(* IEC 61131-3 sources: SortJet_MasterSPS_Aufbau.fbsproj/Device.device.xml.v3^/Plc Logic.plclogic.xml.v3^/Application.application.xml.v3^/09_Station/Stationen/Drehstation [207]/0_Konfig, 3 files *)

(* ---- Antriebsinformationen_207.gvl ---- *)
(* METADATA
{
	"v3Meta": {
		"objectGuid": "9d7b2ddc-bc65-44fc-9f07-0caa3fddbc7e"
	}
}
*)
{attribute 'allow_unqualified_access'}
NAMESPACE Antriebsinformationen_207
VAR_GLOBAL

//-------------------------------------------------------------------------------------------------
// ANTRIEBSINFORMATION [DREHSTATION]
//-------------------------------------------------------------------------------------------------

  apgInfoStation207Glastransport : ARRAY[cWAND_1..cANZAHL_WAENDE] OF AntriebsInformationen := [
    (
      wAchsID                                 :=     17,  // Achs ID aus dem EConSet
      stTyp                                   := 'Belt',  // Typ
      wpSchaltschrank                         :=   2040,  // Daten aus dem Schaltplan
      wpSchaltplanreihe                       :=     02,  // Daten aus dem Schaltplan
      wpSchaltplanseite                       :=    100,  // Daten aus dem Schaltplan
      rpMaxGeschwindigkeit                    :=   1000,  // [mm/s]   Max- Geschwindigkeit für den Automatikbetrieb
      rpHandGeschwindigkeit                   :=    200,  // [mm/s]   Hand- Geschwindigkeit
      rpReduzierteGeschwindigkeit             :=    67,   // [mm/s]   Reduzierte Geschwindigkeit
      rpReferenzGeschwindigkeit               :=      0,  // [mm/s]   Geschwindigkeit für die Referenzfahrt
      rpEinrichtGeschwindigkeit               :=     50,  // [mm/s]   Max Geschwindigkeit während der Einrichtung der Anlage
      rpMaxBeschleunigung                     :=   1500,  // [mm/s^2] Max Beschleunigung
      rpMaxVerzoegerung                       :=   2000,  // [mm/s^2] Max Verzoegerung
      rpMaxRuckzeit                           :=     50,  // [ms]     Ruckzeit des Antriebs
      rpReduzierteBeschleunigung              :=    500,  // [mm/s^2] Reduzierte Beschleunigung
      rpReduzierteVerzoegerung                :=    500,  // [mm/s^2] Reduzierte Verzoegerung
      rpBeschleunigungFremdanlage             :=   1000,  // [mm/s^2] Beschleunigung zu einer Fremdanlage
      rpGeschwindigkeitMessen                 :=    667,  // [mm/s] Geschwindigkeit beim Scheiben messen
      rpGeschwindigkeitSystemcheck            :=  500.0,  // [mm/s]   Geschwindigkeit im Systemcheck (nur Glastransport)
      rpGeschwindigkeitSystemcheckReduzierung :=  167.0,  // [mm/s]   Geschwindigkeit im Systemcheck bei belegtem Vorstop-Sensor (nur Glastransport)
      stOptionen                              := ( eEndschalterQuelle    := Endschalterquelle_EN.KEINE,     // Hardware-Endschalter: KEINE, UMRICHTER oder SPS
                                                   bVersorgungUeberXVR   := FALSE,                          // XVR-Modus: brueckt Hauptschalter 400 V und LS 230 V
                                                   bBremseLoesenFreigabe := FALSE )                         // Der Antrieb darf über eine Betriebsart die Bremse lösen
    )];

  apgInfoStation207GlastransportSlave : ARRAY[cWAND_1..cANZAHL_WAENDE] OF AntriebsInformationen := [
    (
      wAchsID                                 :=     65,  // Achs ID aus dem EConSet
      stTyp                                   := 'Belt',  // Typ
      wpSchaltschrank                         :=   2041,  // Daten aus dem Schaltplan
      wpSchaltplanreihe                       :=     02,  // Daten aus dem Schaltplan
      wpSchaltplanseite                       :=    100,  // Daten aus dem Schaltplan
      rpMaxGeschwindigkeit                    :=      0,  // [mm/s]   Max- Geschwindigkeit für den Automatikbetrieb
      rpHandGeschwindigkeit                   :=      0,  // [mm/s]   Hand- Geschwindigkeit
      rpReduzierteGeschwindigkeit             :=      0,  // [mm/s]   Reduzierte Geschwindigkeit
      rpReferenzGeschwindigkeit               :=      0,  // [mm/s]   Geschwindigkeit für die Referenzfahrt
      rpEinrichtGeschwindigkeit               :=      0,  // [mm/s]   Max Geschwindigkeit während der Einrichtung der Anlage
      rpMaxBeschleunigung                     :=      0,  // [mm/s^2] Max Beschleunigung
      rpMaxVerzoegerung                       :=      0,  // [mm/s^2] Max Verzoegerung
      rpMaxRuckzeit                           :=      0,  // [ms]     Ruckzeit des Antriebs
      rpReduzierteBeschleunigung              :=      0,  // [mm/s^2] Reduzierte Beschleunigung
      rpReduzierteVerzoegerung                :=      0,  // [mm/s^2] Reduzierte Verzoegerung
      rpBeschleunigungFremdanlage             :=      0,  // [mm/s^2] Beschleunigung zu einer Fremdanlage
      rpGeschwindigkeitMessen                 :=      0,  // [mm/s] Geschwindigkeit beim Scheiben messen
      rpGeschwindigkeitSystemcheck            :=  500.0,  // [mm/s]   Geschwindigkeit im Systemcheck (nur Glastransport)
      rpGeschwindigkeitSystemcheckReduzierung :=  167.0,  // [mm/s]   Geschwindigkeit im Systemcheck bei belegtem Vorstop-Sensor (nur Glastransport)
      stOptionen                              := ( eEndschalterQuelle    := Endschalterquelle_EN.KEINE,     // Hardware-Endschalter: KEINE, UMRICHTER oder SPS
                                                   bVersorgungUeberXVR   := FALSE,                          // XVR-Modus: brueckt Hauptschalter 400 V und LS 230 V
                                                   bBremseLoesenFreigabe := FALSE )                         // Der Antrieb darf über eine Betriebsart die Bremse lösen
    )];

  apgInfoStation207Drehen : AntriebsInformationen :=
    (
      wAchsID                                 :=        18,  // Achs ID aus dem EConSet
      stTyp                                   := 'Turning',  // Typ
      wpSchaltschrank                         :=      2042,  // Daten aus dem Schaltplan
      wpSchaltplanreihe                       :=        02,  // Daten aus dem Schaltplan
      wpSchaltplanseite                       :=        65,  // Daten aus dem Schaltplan
      rpMaxGeschwindigkeit                    :=       350,  // [Grad/s] MAX- Geschwindigkeit für die der Antrieb ausgelegt ist // Max 556
      rpHandGeschwindigkeit                   :=       150,  // [Grad/s] Hand- Geschwindigkeit
      rpReduzierteGeschwindigkeit             :=        20,  // [Grad/s] Reduzierte Geschwindigkeit für die bestimmte Situationen
      rpReferenzGeschwindigkeit               :=         1,  // [Grad/s] Geschwindigkeit für die Referenzfahrt
      rpEinrichtGeschwindigkeit               :=        10,  // [Grad/s] Max Geschwindigkeit während der Einrichtung der Anlage
      rpMaxBeschleunigung                     :=       300,  // [Grad/s^2] max Beschleunigung für die der Antrieb ausgelegt ist // Max 1026
      rpMaxVerzoegerung                       :=       300,  // [Grad/s^2] max Verzoegerung für die der Antrieb ausgelegt ist // Max 1026
      rpMaxRuckzeit                           :=       200,   // [ms]     Ruckzeit des Antriebs
      rpReduzierteBeschleunigung              :=       0.5,  // [Grad/s^2] Reduzierte Beschleunigung
      rpReduzierteVerzoegerung                :=       0.5,  // [Grad/s^2] Reduzierte Verzoegerung
      rpBeschleunigungFremdanlage             :=       0.5,  // [Grad/s^2] Beschleunigung zu einer Fremd-Anlage
      rpGeschwindigkeitMessen                 :=         0,  // [Grad/s] Geschwindigkeit für die Messfahrt
      rpGeschwindigkeitSystemcheck            :=  500.0,  // [mm/s]   Geschwindigkeit im Systemcheck (nur Glastransport)
      rpGeschwindigkeitSystemcheckReduzierung :=  167.0,  // [mm/s]   Geschwindigkeit im Systemcheck bei belegtem Vorstop-Sensor (nur Glastransport)
      stOptionen                              := ( eEndschalterQuelle    := Endschalterquelle_EN.UMRICHTER, // Hardware-Endschalter: KEINE, UMRICHTER oder SPS
                                                   bVersorgungUeberXVR   := FALSE,                          // XVR-Modus: brueckt Hauptschalter 400 V und LS 230 V
                                                   bBremseLoesenFreigabe := FALSE )                         // Der Antrieb darf über eine Betriebsart die Bremse lösen
    );

  apgInfoStation207Kippen : AntriebsInformationen :=
    (
      wAchsID                                 :=        65,  // Achs ID aus dem EConSet
      stTyp                                   := 'Tilting',  // Typ
      wpSchaltschrank                         :=      2043,  // Daten aus dem Schaltplan
      wpSchaltplanreihe                       :=         2,  // Daten aus dem Schaltplan
      wpSchaltplanseite                       :=       100,  // Daten aus dem Schaltplan
      rpMaxGeschwindigkeit                    :=      1400,  // [Grad/s] Max- Geschwindigkeit für die der Antrieb ausgelegt ist
      rpHandGeschwindigkeit                   :=      1400,  // [Grad/s] Hand- Geschwindigkeit
      rpReduzierteGeschwindigkeit             :=       800,  // [Grad/s] Reduzierte Geschwindigkeit für die bestimmte Situationen
      rpReferenzGeschwindigkeit               :=       100,  // [Grad/s] Geschwindigkeit für die Referenzfahrt
      rpEinrichtGeschwindigkeit               :=       100,  // [Grad/s] Max Geschwindigkeit während der Einrichtung der Anlage
      rpMaxBeschleunigung                     :=       250,  // [Grad/s^2] Max Beschleunigung für die der Antrieb ausgelegt ist
      rpMaxVerzoegerung                       :=       250,  // [Grad/s^2] Max Verzoegerung für die der Antrieb ausgelegt ist
      rpMaxRuckzeit                           :=        50,  // [ms] Ruckzeit des Antriebs
      rpReduzierteBeschleunigung              :=       100,  // [Grad/s^2] Reduzierte Beschleunigung
      rpReduzierteVerzoegerung                :=       100,  // [Grad/s^2] Reduzierte Verzoegerung
      rpBeschleunigungFremdanlage             :=         1,  // [Grad/s^2] Beschleunigung zu einer Fremd-Anlage
      rpGeschwindigkeitMessen                 :=         0,  // [Grad/s] Geschwindigkeit für die Messfahrt
      rpGeschwindigkeitSystemcheck            := 500.0,  // [mm/s]   Geschwindigkeit im Systemcheck (nur Glastransport)
      rpGeschwindigkeitSystemcheckReduzierung := 167.0,  // [mm/s]   Geschwindigkeit im Systemcheck bei belegtem Vorstop-Sensor (nur Glastransport)
      stOptionen                              := ( eEndschalterQuelle    := Endschalterquelle_EN.UMRICHTER, // Hardware-Endschalter: KEINE, UMRICHTER oder SPS
                                                   bVersorgungUeberXVR   := FALSE,                          // XVR-Modus: brueckt Hauptschalter 400 V und LS 230 V
                                                   bBremseLoesenFreigabe := FALSE )                         // Der Antrieb darf über eine Betriebsart die Bremse lösen
    );

    apgInfoStation207Querfahrt : AntriebsInformationen :=
    (
      wAchsID                                 :=         65,  // Achs ID aus dem EConSet
      stTyp                                   := 'Movement',  // Typ
      wpSchaltschrank                         :=       2044,  // Daten aus dem Schaltplan
      wpSchaltplanreihe                       :=         02,  // Daten aus dem Schaltplan
      wpSchaltplanseite                       :=        100,  // Daten aus dem Schaltplan
      rpMaxGeschwindigkeit                    :=        250,  // [mm/s] MAX- Geschwindigkeit für die der Antrieb ausgelegt ist
      rpHandGeschwindigkeit                   :=        100,  // [mm/s] Hand- Geschwindigkeit
      rpReduzierteGeschwindigkeit             :=         50,  // [mm/s] Reduzierte Geschwindigkeit für die bestimmte Situationen
      rpReferenzGeschwindigkeit               :=         20,  // [mm/s] Geschwindigkeit für die Referenzfahrt
      rpEinrichtGeschwindigkeit               :=         50,  // [mm/s] Max Geschwindigkeit während der Einrichtung der Anlage
      rpMaxBeschleunigung                     :=        600,  // [mm/s^2] max Beschleunigung für die der Antrieb ausgelegt ist
      rpMaxVerzoegerung                       :=        600,  // [mm/s^2] max Verzoegerung für die der Antrieb ausgelegt ist
      rpMaxRuckzeit                           :=        600,  // [ms]     Ruckzeit des Antriebs
      rpReduzierteBeschleunigung              :=        200,  // [mm/s^2] Reduzierte Beschleunigung
      rpReduzierteVerzoegerung                :=        200,  // [mm/s^2] Reduzierte Verzoegerung
      rpBeschleunigungFremdanlage             :=          0,  // [mm/s^2] Beschleunigung zu einer Fremd-Anlage
      rpGeschwindigkeitMessen                 :=          0,  // [mm/s] Geschwindigkeit für die Messfahrt
      rpGeschwindigkeitSystemcheck            := 500.0,  // [mm/s]   Geschwindigkeit im Systemcheck (nur Glastransport)
      rpGeschwindigkeitSystemcheckReduzierung := 167.0,  // [mm/s]   Geschwindigkeit im Systemcheck bei belegtem Vorstop-Sensor (nur Glastransport)
      stOptionen                              := ( eEndschalterQuelle    := Endschalterquelle_EN.UMRICHTER, // Hardware-Endschalter: KEINE, UMRICHTER oder SPS
                                                   bVersorgungUeberXVR   := FALSE,                          // XVR-Modus: brueckt Hauptschalter 400 V und LS 230 V
                                                   bBremseLoesenFreigabe := FALSE )                         // Der Antrieb darf über eine Betriebsart die Bremse lösen
    );

END_VAR

END_NAMESPACE

(* ---- MK_Station_207.gvl ---- *)
(* METADATA
{
	"v3Meta": {
		"objectGuid": "ad0b4350-ba92-412a-9245-7792853cbecb"
	}
}
*)
{attribute 'allow_unqualified_access'}
NAMESPACE MK_Station_207
VAR_GLOBAL

//-------------------------------------------------------------------------------------------------
// MASCHINEPARAMETER: DREHSTATION
//-------------------------------------------------------------------------------------------------

  apgMKStation207 : Parameter_Station:=
    (
      stStationsNummern                     := ( NummerIntern :=   207,                                                      // Stationsnummer fuer das MMI und die Stationsangabe der Meldungen
                                                 NummerExtern :=  1207,                                                      // Stationsnummer fuer Bedienermeldungen
                                                 NummerSPS    :=   207 ),                                                    // Stationsnummer SPS-intern (Indizes)
      bDeaktivieren                         := FALSE,                                                                        // Station deaktiviert (keine Auftraege, keine Referenzfahrt)
      wMeldungsNummer                       := 1810,                                                                         // Basis-Meldungsnummer (WatchIO)
      eStationsTyp                          := eStation,                                                                     // Typ der Station
      eaAutomatikkreis                      := [eAutomatikkreis_1],                                                          // Automatikkreise, zu denen die Station gehoert
      eaSicherheitskreis                    := [eSicherheitskreis_1, eSicherheitskreis_4],                                   // Sicherheitskreise, in die die Station eingebunden ist
      astSicherheitskreisTeilabschaltung    := [ ( eSicherheitskreis := eSicherheitskreis_4,                                 // SK4 (Abschrankung 208) schaltet nur Drehen/Kippen ab,
                                                   bTeilabschaltung  := TRUE,                                                //   Glastransport, Geblaese, Querfahrt und Pneumatik bleiben aktiv
                                                   bDrehen           := TRUE,
                                                   bKippen           := TRUE ) ],
      eSystemcheckZyklus                    := eSystemcheckZyklus_1,                                                         // In welchem Zyklus des Systemchecks die Station geprueft wird
      stSchnittstellendaten                 := ( wVorgaengerStation := cSTATION_DYNAMISCH,                                   // Station vor dieser Station (cSTATION_DYNAMISCH bei mehreren)
                                                 wNachfolgerStation := cSTATION_DYNAMISCH,                                   // Station nach dieser Station (cSTATION_DYNAMISCH bei mehreren)
                                                 bStationIstShuttle := FALSE                                                 // Station ist ein Shuttle
                                               ),
      stStationsOptionen                    := ( stSystemcheck :=  ( bScheibenVermessenSystemCheck               := TRUE,    // Scheiben im Systemcheck vermessen
                                                                     bScheibeNachSystemcheckAufAuslauf           := TRUE,    // Scheibe nach dem Systemcheck auf den Auslaufsensor fahren
                                                                     bSystemCheckMitVorgaengerBatchTransport     := FALSE,   // derzeit ohne Funktion
                                                                     bSystemCheckMitNachfolgerBatchTransport     := FALSE,   // derzeit ohne Funktion
                                                                     bOptionSystemCheckScheibeMittigLegen        := FALSE ), // derzeit ohne Funktion

                                                 // stTransfershuttle
                                                 stGlastransport :=  ( bVortransport                             := FALSE,   // Vortransport aktivieren [Bsp.: Nach einem Eintransport mit gesetztem Bit <Letzte Scheibe>]
                                                                       bTransportMasterSlaveEintransport         := FALSE,   // derzeit ohne Funktion
                                                                       bTransportMasterSlaveAustransport         := TRUE ,   // Austransport als Slave auf die Achse des Nachfolgers
                                                                       bGLasUebernahmeSenkrecht                  := FALSE,   // RKT - Eintransport in Senkrechter-Position bzw. in Waagerechter- Position [default]
                                                                       bAustransportISOLinie                     := FALSE,   // Austransport an eine ISO-Linie
                                                                       bScheibenVermessen                        := FALSE,   // Scheibenmessung am Anlegetisch/Anlegewand
                                                                       bMessrichtungNegativ                      := FALSE,   // Negative Fahrtrichtung beim Messen
                                                                       bScheibenmessungEintransport              := FALSE,   // Scheibenmessung beim Eintransport
                                                                       bScheibenmessungSensorVorabAuslauf        := FALSE    // Scheibenmessung mit SensorVorabAuslauf z.B. Anlegewand
                                                                      ),
                                                 // stAnlegetisch
                                                 // stEckuebergabe
                                                 stDrehstation   :=  ( bDrehpositionenVomMMI                     := FALSE,            // TRUE: Drehpositionen aus den MMI-Auftragsdaten; FALSE: aus der Stationskonfiguration [aEintransporte/aAustransporte]
                                                                       wStandardTransferstation                  := cSTATION_206 ),   // Systemcheck (Drehpositionen nicht vom MMI): Transferstation, wenn die Auftragsdaten 0 enthalten
                                                 bVorAbKomponentenAnsteuerung              := FALSE,                         // VorAbKomponentenAnsteuerung Auftraege werden bearbeitet
                                                 bVerstellungEinAusGefahrenLogikDrehen     := FALSE,                         // Verstellung: Logik ein-/ausgefahren gedreht
                                                 bLangsamfahrtNockenQuerfahrtAktivieren    := FALSE,                         // Querfahrt: Langsamfahrt-Nocken auswerten
                                                 bSKBlockierenDurchVorabSensoren           := FALSE,                         // Vorab-Sensoren belegt blockieren das Oeffnen des Sicherheitskreises
                                                 bStationLeerfahrenBeiSkAnforderung        := FALSE,                         // Station bei Anforderung Sicherheitskreis leerfahren
                                                 bGlasAbgenommenAutomatischQuittieren      := FALSE,                         // derzeit ohne Funktion
                                                 bScheibeAbnehmenNachEintransport          := FALSE                          // Scheibe nach dem Eintransport wieder abnehmen
                                               ),
      stStationsAufbau                      := ( bGeblase                      := [ cANZAHL_WAENDE(TRUE) ],                  // Ausbaustufe: Geblaese je Wand
                                                 bGlastransport                := [ cANZAHL_WAENDE(TRUE) ],                  // Ausbaustufe: Glastransport je Wand
                                                 bKippen                       := [ cANZAHL_WAENDE(TRUE) ],                  // Ausbaustufe: Kippen je Wand
                                                 bKippenSchuetz                := TRUE,                                      // Kippen ueber Schuetz statt Umrichter
                                                 bTransportVerstellung         := [ cANZAHL_WAENDE(FALSE) ],                 // Ausbaustufe Shuttle: Transport-/Dickenverstellung je Wand
                                                 bHub                          := FALSE,                                     // Ausbaustufe: Hub der Station
                                                 bHubrahmen                    := FALSE,                                     // Ausbaustufe: Hubrahmen (Riemen heben/senken)
                                                 bDrehen                       := TRUE,                                      // Ausbaustufe: Drehen
                                                 bQuerachse                    := FALSE,                                     // Ausbaustufe: Querachse
                                                 bMessachse                    := FALSE,                                     // Ausbaustufe: Messachse (Anlegetisch, Anlegewand)
                                                 bDruckluft                    := TRUE,                                      // Druckluftueberwachung vorhanden
                                                 bAnschlag                     := FALSE,                                     // Ausbaustufe: Ausrichtanschlaege
                                                 bSensorAuslauf                := TRUE,                                      // Auslaufsensor vorhanden
                                                 bSensorEinlauf                := TRUE,                                      // Einlaufsensor vorhanden
                                                 bSensorEinlaufStopp           := FALSE,                                     // Shuttle: zusaetzlicher Stopp-Sensor am Einlauf (ohne: Einlaufsensor), Gegenstueck zum Auslauf-Stopp im Rueckwaertstransport
                                                 bSensorAuslaufStopp           := FALSE,                                     // Shuttle: zusaetzlicher Stopp-Sensor am Auslauf (ohne: Auslaufsensor), Verfahrfreigabe und Scheibe hat Shuttle verlassen
                                                 bDurchlaufSperreZumNachfolger := FALSE,                                     // Ausbaustufe: bewegliche Abschrankung zum Nachfolger
                                                 bQuerfahrt                    := FALSE,                                     // Ausbaustufe: Querfahrt
                                                 bKipparme                     := FALSE,                                     // Ausbaustufe: Kipparme
                                                 bSlaveAntrieb                 := FALSE,                                     // Glastransport mit Slave-Antrieb
                                                 bMessachseAmEndeVomTisch      := FALSE,                                     // Messachse am Ende des Tisches (Hoehenfehler fragt den Bediener)
                                                 bWandverstellung              := [ FALSE ],                                 // Ausbaustufe Station: Wandverstellung je Wand
                                                 bWandverstellungMotorisch     := FALSE,                                     // Shuttle: Transport-/Wandverstellung mit Antrieb statt pneumatisch
                                                 bRoellchenleiste              := [ FALSE ],                                 // Ausbaustufe Station: Roellchenleiste je Wand
                                                 bDurchgang                    := FALSE,                                     // Station ist Teil eines Durchgangs (belegt = Oeffnen blockiert)
                                                 bRolltor                      := FALSE,                                     // Ausbaustufe Faecherwagen: Rolltor
                                                 bKlemmzylinder                := FALSE,                                     // Ausbaustufe Faecherwagen: Klemmzylinder fixiert den Oberrahmen beim Ein- und Ausschleusen
                                                 bGreifer                      := [cANZAHL_WAENDE(FALSE)],                   // Shuttle: Greifer je Wand (Scheibe aus dem Faecherwagen ziehen bzw. hineinschieben)
                                                 bRFID                         := FALSE,                                     // RFID-Leser vorhanden
                                                 bAGV                          := FALSE,                                     // Ausbaustufe Faecherwagen: Betrieb mit AGV
                                                 bDLSSchmiersystem             := FALSE,                                     // Zentralschmierung DLS vorhanden
                                                 bGlastransportSlaveVorhanden  := FALSE,                                     // Glastransport mit Slave-Antrieb (Meldungen/Ueberwachung Slave)
                                                 wHydraulikstation             := 0                                          // Faecherwagen Hydraulik: zugeordnete Hydraulikstation (cHYDRAULIKSTATION_x), 0 = keine
                                               ),
      stStationsParameter                   := ( rLaengeUebergroesseScheibe              := 4240,                            // Shuttle: ab dieser Scheibenlaenge gilt die Scheibe als uebergross [mm]
                                                 rMinGlasHoeheAutomatischenEintransport  := 500,                             // VSG: Mindesthoehe fuer automatischen Eintransport [mm]
                                                 rMinGlasLaengeAutomatischenEintransport := 500,                             // VSG: Mindestlaenge fuer automatischen Eintransport [mm]
                                                 wMaximaleAnzahlAktiverAuftraege := 1,                                       // derzeit ohne Funktion
                                                 rMinPosSwEsEingrenzung                  := 0.0,                             // Externer zusaetzlicher Software-Endschalter MIN; 0 = inaktiv; darf den MK-MIN nur weiter eingrenzen
                                                 rMaxPosSwEsEingrenzung                  := 0.0,                             // Externer zusaetzlicher Software-Endschalter MAX; 0 = inaktiv; darf den MK-MAX nur weiter eingrenzen
                                                 rPosFreigabePufferAusfahren             := 0.0                              // derzeit ohne Funktion
                                              ),
      // stFremdanlage
      stGlasdaten                           := [(
                                                 rlMinGlasLaenge                  := 350,                                    // minimal zulässige GlasLänge
                                                 rlMaxGlasLaenge                  := 2500,                                   // maximale zulässige GlasLänge
                                                 rlMinGlasHoehe                   := 190,                                    // minimal zulässige GlasHöhe
                                                 rlMaxGlasHoehe                   := 1800,                                   // maximale zulässige GlasHöhe
                                                 rlMinGlasDicke                  := 3,                                     // minimal zulässige GlasDicke
                                                 rlMaxGlasDicke                  := 12.76,                                      // maximal zulaessige Glasdicke [mm]
                                                 rlLaengeMaxGlas                  := 0.0                                     // maximal zulaessige Glaslaenge [mm]
                                               )]
      // astShuttleAnhaltenQuellen
    );

  apgMKStation207Glastransport : ARRAY[cWAND_1..cANZAHL_WAENDE] OF Parameter_Glastransport := [
    (
      rLaengeStation                        := 2800, // Länge der Station
      rScheibenabstand                      :=  300, // Der Abstand zwischen zwei Scheiben auf der Station
      rWegUeberAuslauf                      :=   50, // Weg ueber den Auslaufsensor hinaus [mm]
      rWegUeberEinlauf                      :=   50, // Weg ueber den Einlaufsensor hinaus [mm]
      rWegUeberSensorenSystemCheck          :=   15, // Der Weg der Ueber ein die Sensoren zum vermessen der Scheiben
      rUeberwachungAuslaufsensor            :=  500, // Ueberwachung des Auslaufsensors [Strecke in der der Auslaufsensor Frei / ueberfahren werden soll]
      rUeberwachungEinlaufsensor            :=  500, // Ueberwachung des Einlaufsensors [Strecke in der der Einlaufsensor Frei / ueberfahren werden soll]
      rWegUeberEinlaufEintransport          :=  150, // Eintransport vorwaerts: Abstand Scheibenhinterkante zum Einlaufsensor [mm]
      rWegUeberEinlaufAustransport          :=   50, // Lage Auf Einlauf: Scheibe liegt um diesen Weg auf dem Einlaufsensor [mm]
      rWegUeberAuslaufEintransport          :=   50, // Eintransport rueckwaerts: Abstand Scheibenhinterkante zum Auslaufsensor [mm]
      rWegUeberAuslaufAustransport          :=   10, // Lage Auf Auslauf: Weg ueber den Auslaufsensor hinaus [mm]
      rWegEinlaufsensorZuVorStopSensor      := 2700, // Beschreibt den Weg vum eine Scheibe beim EIntransport vom Einlaufsensor bis ueberden Vorabstopsensor zu verfahren
      rMesstoleranz                         :=   10, // Toleranz-Mass fuer die Scheibenlaengenmessung
      rMessstrecke                          := 2740, // Beschreibt die Strecke ziwischen 2 Sensoren die der Antrieb verfaehrt
      rWegstreckeBisZurVerzoegerung         := 2200  // Beschreibt die Strecke die gefahren werden soll bis der Antrieb abgebremst werden soll, dies gilt fuer Eintransportauftraege die das Bit "Letzte Scheibe" gesetzt haben
    )];

  apgMKStation207Drehen : Parameter_Drehen :=
    (
      tZeitAntriebsfreigabeErhalten        := T#180S,               // [ms \ s] Energieeinsparrung: Zeiteinheit nach der die Antriebsfreigabe entzogen werden soll wenn keine Aktion ansteht [1 s = 1000 ms ]
      rToleranz                            :=    0.1,               // Toleranz beim Entscheiden der aktuellen Position
      rDrehposition_0_Grad                 := 880.87,               // Drehposition fuer die 0 Grad   -> Shuttle 101 / Kipptisch 206 (bisher 90 Grad)
      rDrehposition_90_Grad                :=    441,               // Drehposition fuer die 90 Grad  -> Anlegewand 208 (bisher 0 Grad)
      rDrehposition_180_Grad               :=   2.83,               // Drehposition fuer die 180 Grad -> Shuttle 101 / Kipptisch 206 (gedreht)
      rDrehposition_270_Grad               :=      0,               // Drehposition fuer die 270 Grad
      bArretierung                         :=    TRUE,              // Arretierung vorhanden
      eZielDrehpositionLeer                := eDrehPosition0Grad,   // derzeit ohne Funktion
      astKippenJeDrehposition              := [ ( eKippenOhneLetzteScheibe := eKippen_Position_84Grad,     // [0]   0 Grad -> Shuttle 101 / Kipptisch 206 (TODO: ohne letzte Scheibe 90 Grad, sobald der RKT auf 90 Grad kippt und die Drehpositionen vom MMI kommen)
                                                  eKippenMitLetzterScheibe := eKippen_Position_90Grad ),
                                                ( eKippenOhneLetzteScheibe := eKippen_Position_84Grad,     // [1]  90 Grad -> Anlegewand 208
                                                  eKippenMitLetzterScheibe := eKippen_Position_84Grad ),
                                                ( eKippenOhneLetzteScheibe := eKippen_Position_84Grad,     // [2] 180 Grad -> Shuttle 101 / Kipptisch 206 (TODO: ohne letzte Scheibe 90 Grad, sobald der RKT auf 90 Grad kippt und die Drehpositionen vom MMI kommen)
                                                  eKippenMitLetzterScheibe := eKippen_Position_90Grad ),
                                                ( eKippenOhneLetzteScheibe := eKippen_Default,             // [3] 270 Grad -> nicht genutzt
                                                  eKippenMitLetzterScheibe := eKippen_Default ) ]
    );

  apgMKStation207Kippen : ARRAY[cWAND_1..cANZAHL_WAENDE] OF Parameter_Kippen := [
    (
       tZeitlicheUeberwachungKippen          :=  T#30S, // [ms \ s] Verwendet fuer Antriebe die Ueber einen Schuetz angesteuert werden
       tZeitAntriebsfreigabeErhalten         := T#100S, // [ms \ s] Energieeinsparrung: Zeiteinheit nach der die Antriebsfreigabe entzogen werden soll wenn keine Aktion ansteht [1 s = 1000 ms ]
       rToleranz                             :=      2, // Toleranz beim Entscheiden der aktuellen Position
       rPosition0Grad                        :=      0, // Waagerechte- Position 0 Grad: Position auf die die Station gehoben werden soll
       rPosition84Grad                       :=      0, // Senkrechte- Position 84 Grad: Position auf die die Station gehoben werden soll
       rPosition90Grad                       :=      0, // Senkrechte-Position 90 Grad : Position auf die die Station gesenkt werden soll
       rPosition96Grad                       :=      0, // Senkrechte-Position 96 Grad : Position auf die die Station gesenkt werden soll
       bKippenMitSchuetz                     :=  TRUE,  // Kippen per Umrichter oder Schütz
       rPosition88_5Grad                     := 0.0     // Senkrechte- Position 84 Grad: Position auf die die Station gehoben werden soll
    )];

  apgMKStation207Querfahrt : Parameter_Querfahrt :=
    (
      tZeitAntriebsfreigabeErhalten          := T#10S // Energieeinsparung: Zeit nach der die Antriebsfreigabe entzogen wird, wenn keine Aktion ansteht
    );

END_VAR
END_NAMESPACE

(* ---- Konfiguration_207.gvl ---- *)
(* METADATA
{
	"v3Meta": {
		"objectGuid": "07d733b1-5f14-4340-93e0-09bebec56eed"
	}
}
*)
{attribute 'allow_unqualified_access'}
NAMESPACE Konfiguration_207
VAR_CONFIG

  // GEBLÄSE
  Globale_Bausteine.Drehstation207.Geblaese.in_bMotorschutzschalter_OK                      AT %MX1.1   : BOOL; // OPTION
  Globale_Bausteine.Drehstation207.Geblaese.out_bStarteGeblaese                             AT %MX2071.2 : BOOL; // OPTION

  // KIPPEN
  Globale_Bausteine.Drehstation207.Kippen.in_bMotorschutzschalter_OK                        AT %IX1.7   : BOOL; // IO-L - 207 kippen Motorstarter / Sicherung OK
  Globale_Bausteine.Drehstation207.Kippen.in_bMotorstarter_OK                               AT %MX1.1   : BOOL; // OPTION
  Globale_Bausteine.Drehstation207.Kippen.in_bLSBremse_OK                                   AT %MX1.1   : BOOL; // OPTION
  Globale_Bausteine.Drehstation207.Kippen.in_bLS400V_OK                                     AT %MX1.1   : BOOL; // OPTION

  Globale_Bausteine.Drehstation207.Kippen.out_bKippen84Grad                                 AT %QX1.2   : BOOL; // IO-L - 207 kippen 1 nach 84 Grad
  Globale_Bausteine.Drehstation207.Kippen.out_bKippen90Grad                                 AT %QX1.1   : BOOL; // IO-L - 207 kippen 1 nach 90 Grad
  Globale_Bausteine.Drehstation207.Kippen.out_bBremseLoesen                                 AT %MX2070.0 : BOOL; // OPTION
  Globale_Bausteine.Drehstation207.Kippen.out_bReset                                        AT %MX2070.1 : BOOL; // OPTION

  // WANDVERSTELLUNG
  Globale_Bausteine.Drehstation207.Dickenverstellung.in_bStatusZylinder1Ausgefahren         AT %MX1.0   : BOOL; // OPTION
  Globale_Bausteine.Drehstation207.Dickenverstellung.in_bStatusZylinder1Eingefahren         AT %MX1.0   : BOOL; // OPTION
  Globale_Bausteine.Drehstation207.Dickenverstellung.in_bStatusZylinder2Ausgefahren         AT %MX1.0   : BOOL; // OPTION
  Globale_Bausteine.Drehstation207.Dickenverstellung.in_bStatusZylinder2Eingefahren         AT %MX1.0   : BOOL; // OPTION

  Globale_Bausteine.Drehstation207.Dickenverstellung.out_bZylinder1Ausfahren                AT %MX2071.0 : BOOL; // OPTION
  Globale_Bausteine.Drehstation207.Dickenverstellung.out_bZylinder1Einfahren                AT %MX2071.1 : BOOL; // OPTION
  Globale_Bausteine.Drehstation207.Dickenverstellung.out_bZylinder2Ausfahren                AT %MX2070.2 : BOOL; // OPTION
  Globale_Bausteine.Drehstation207.Dickenverstellung.out_bZylinder2Einfahren                AT %MX2070.3 : BOOL; // OPTION

  // QUERACHSE
  Globale_Bausteine.Drehstation207.Querachse.in_bStatusZylinder1Ausgefahren                AT %MX1.0   : BOOL; // OPTION
  Globale_Bausteine.Drehstation207.Querachse.in_bStatusZylinder1Eingefahren                AT %MX1.0   : BOOL; // OPTION
  Globale_Bausteine.Drehstation207.Querachse.in_bStatusZylinder2Ausgefahren                AT %MX1.0   : BOOL; // OPTION
  Globale_Bausteine.Drehstation207.Querachse.in_bStatusZylinder2Eingefahren                AT %MX1.0   : BOOL; // OPTION

  Globale_Bausteine.Drehstation207.Querachse.out_bZylinder1Ausfahren                       AT %MX2070.4 : BOOL; // OPTION
  Globale_Bausteine.Drehstation207.Querachse.out_bZylinder1Einfahren                       AT %MX2070.5 : BOOL; // OPTION
  Globale_Bausteine.Drehstation207.Querachse.out_bZylinder2Ausfahren                       AT %MX2070.6 : BOOL; // OPTION
  Globale_Bausteine.Drehstation207.Querachse.out_bZylinder2Einfahren                       AT %MX2070.7 : BOOL; // OPTION

END_VAR

END_NAMESPACE
